(* IEC 61131-3 sources: rusty/tests/lit/cfc/validation/function_inout_negated, 2 files *)

(* ---- addInto.st ---- *)
FUNCTION addInto : DINT
VAR_INPUT
    delta : DINT;
END_VAR
VAR_IN_OUT
    acc : DINT;
END_VAR
    acc := acc + delta;
    addInto := acc;
END_FUNCTION

(* ---- main.st ---- *)
// A negated inout pin transpiles like an input pin, but an inout passes by
// reference and a NOT expression has no storage behind it, so validation
// rejects the call.
// CHECK: {{.*}}function_inout_negated.cfc.function_inout_negated:1:1: error[E031]: Expected a reference for parameter acc because their type is InOut
// CHECK: error: Compilation aborted due to critical errors
FUNCTION main : DINT
END_FUNCTION
